INTERFACE I_Logger

METHOD Log : BOOL
VAR_INPUT
  sMessage  : STRING;
  nSeverity  : INT;
END_VAR
END_METHOD

END_INTERFACE

(* stored: Version 1.1.0.1, ProductVersion 3.1.4024.12
   Itf I_Logger: Id {0a1b2c3d-0000-4000-8000-000000000002}
   Method Log: Id {0a1b2c3d-0000-4000-8000-000000000003} *)
